Fanuc KAREL source: KT00846.KL

PROGRAM KT00846
%NOLOCKGROUP
VAR
  R1: REAL
  R2: REAL
  OUT: INTEGER
BEGIN
  R1 = 2.0
  R2 = 3.0
  R1 = 2.0
  R2 = 3.0
  OUT = TAN(R1)
END KT00846
